TYPE "DT_ALM_SYSTEM_SPARE_26"
VERSION : 0.1
   STRUCT
      LINE_2_DS_ERR { S7_SetPoint := 'False'} : "DT_ALM_SOLO" := (832, FALSE, FALSE, TRUE, (), (), 6, 0, 4, (), (), (), (), (), T#50MS);
      LINE_2_DS_OFF { S7_SetPoint := 'False'} : "DT_ALM_SOLO" := (833, FALSE, FALSE, TRUE, (), (), 6, 0, 4, (), (), (), (), (), T#50MS);
      LINE_2_DS_GND { S7_SetPoint := 'False'} : "DT_ALM_SOLO" := (834, FALSE, FALSE, FALSE, (), (), 0, 0, 0, (), (), (), (), (), T#500MS);
      LINE_2_ES_ERR { S7_SetPoint := 'False'} : "DT_ALM_SOLO" := (835, FALSE, FALSE, TRUE, (), (), 6, 0, 4, (), (), (), (), (), T#50MS);
      LINE_2_ES_OFF { S7_SetPoint := 'False'} : "DT_ALM_SOLO" := (836, FALSE, FALSE, FALSE, (), (), 0, 0, 0, (), (), (), (), (), T#500MS);
      LINE_2_ES_GND { S7_SetPoint := 'False'} : "DT_ALM_SOLO" := (837, FALSE, FALSE, TRUE, (), (), 6, 0, 4, (), (), (), (), (), T#50MS);
      LINE_2_NO_VOLTAGE { S7_SetPoint := 'False'} : "DT_ALM_SOLO" := (838, FALSE, FALSE, TRUE, (), (), 6, 0, 4, (), (), (), (), (), T#50MS);
      LINE_2_SYNCH_VT_MCB_OFF { S7_SetPoint := 'False'} : "DT_ALM_SOLO" := (839, FALSE, FALSE, FALSE, (), (), 0, 0, 0, (), (), (), (), (), T#500MS);
      LINE_2_CB_SPRING { S7_SetPoint := 'False'} : "DT_ALM_SOLO" := (840, FALSE, FALSE, TRUE, (), (), 6, 0, 1, (), (), (), (), (), T#50MS);
      LINE_2_CB_UNLOCKED { S7_SetPoint := 'False'} : "DT_ALM_SOLO" := (841, FALSE, FALSE, FALSE, (), (), 0, 0, 0, (), (), (), (), (), T#500MS);
      LINE_2_CB_LOCAL { S7_SetPoint := 'False'} : "DT_ALM_SOLO" := (842, FALSE, FALSE, FALSE, (), (), 0, 0, 0, (), (), (), (), (), T#500MS);
      LINE_2_CB_ERR { S7_SetPoint := 'False'} : "DT_ALM_SOLO" := (843, FALSE, FALSE, TRUE, (), (), 6, 0, 4, (), (), (), (), (), T#50MS);
      LINE_2_CB_OFF { S7_SetPoint := 'False'} : "DT_ALM_SOLO" := (844, FALSE, FALSE, TRUE, (), (), 6, 0, 4, (), (), (), (), (), T#50MS);
      LINE_2_CB_APU_ERR { S7_SetPoint := 'False'} : "DT_ALM_SOLO" := (845, FALSE, FALSE, FALSE, (), (), 0, 0, 0, (), (), (), (), (), T#500MS);
      LINE_2_MCB_W { S7_SetPoint := 'False'} : "DT_ALM_SOLO" := (846, FALSE, FALSE, FALSE, (), (), 0, 0, 0, (), (), (), (), (), T#500MS);
      LINE_2_MCB_T { S7_SetPoint := 'False'} : "DT_ALM_SOLO" := (847, FALSE, FALSE, TRUE, (), (), 6, 0, 4, (), (), (), (), (), T#50MS);
      LINE_2_CNTRL_MCB_OFF { S7_SetPoint := 'False'} : "DT_ALM_SOLO" := (848, FALSE, FALSE, FALSE, (), (), 0, 0, 0, (), (), (), (), (), T#500MS);
      LINE_2_MCBS_ALARM { S7_SetPoint := 'False'} : "DT_ALM_SOLO" := (849, FALSE, FALSE, FALSE, (), (), 0, 0, 0, (), (), (), (), (), T#500MS);
      LINE_2_MCBS_TRIP { S7_SetPoint := 'False'} : "DT_ALM_SOLO" := (850, FALSE, FALSE, FALSE, (), (), 0, 0, 0, (), (), (), (), (), T#500MS);
      SPARE_819 { S7_SetPoint := 'False'} : "DT_ALM_SOLO" := (851, FALSE, FALSE, FALSE, (), (), 0, 0, 0, (), (), (), (), (), T#500MS);
      SPARE_820 { S7_SetPoint := 'False'} : "DT_ALM_SOLO" := (852, FALSE, FALSE, FALSE, (), (), 0, 0, 0, (), (), (), (), (), T#500MS);
      SPARE_821 { S7_SetPoint := 'False'} : "DT_ALM_SOLO" := (853, FALSE, FALSE, FALSE, (), (), 0, 0, 0, (), (), (), (), (), T#500MS);
      SPARE_822 { S7_SetPoint := 'False'} : "DT_ALM_SOLO" := (854, FALSE, FALSE, FALSE, (), (), 0, 0, 0, (), (), (), (), (), T#500MS);
      SPARE_823 { S7_SetPoint := 'False'} : "DT_ALM_SOLO" := (855, FALSE, FALSE, FALSE, (), (), 0, 0, 0, (), (), (), (), (), T#500MS);
      SPARE_824 { S7_SetPoint := 'False'} : "DT_ALM_SOLO" := (856, FALSE, FALSE, FALSE, (), (), 0, 0, 0, (), (), (), (), (), T#500MS);
      SPARE_825 { S7_SetPoint := 'False'} : "DT_ALM_SOLO" := (857, FALSE, FALSE, FALSE, (), (), 0, 0, 0, (), (), (), (), (), T#500MS);
      SPARE_826 { S7_SetPoint := 'False'} : "DT_ALM_SOLO" := (858, FALSE, FALSE, FALSE, (), (), 0, 0, 0, (), (), (), (), (), T#500MS);
      SPARE_827 { S7_SetPoint := 'False'} : "DT_ALM_SOLO" := (859, FALSE, FALSE, FALSE, (), (), 0, 0, 0, (), (), (), (), (), T#500MS);
      SPARE_828 { S7_SetPoint := 'False'} : "DT_ALM_SOLO" := (860, FALSE, FALSE, FALSE, (), (), 0, 0, 0, (), (), (), (), (), T#500MS);
      SPARE_829 { S7_SetPoint := 'False'} : "DT_ALM_SOLO" := (861, FALSE, FALSE, FALSE, (), (), 0, 0, 0, (), (), (), (), (), T#500MS);
      SPARE_830 { S7_SetPoint := 'False'} : "DT_ALM_SOLO" := (862, FALSE, FALSE, FALSE, (), (), 0, 0, 0, (), (), (), (), (), T#500MS);
      SPARE_831 { S7_SetPoint := 'False'} : "DT_ALM_SOLO" := (863, FALSE, FALSE, FALSE, (), (), 0, 0, 0, (), (), (), (), (), T#500MS);
   END_STRUCT;

END_TYPE

